Fanuc KAREL source: KT00497.KL

PROGRAM KT00497
%NOLOCKGROUP
VAR
  P1: XYZWPR
  P2: POSITION
  OUT: JOINTPOS
BEGIN
  P1.X = 1.0
  OUT = P1 : P2
END KT00497
